Fanuc KAREL source: kt00161.KL

-- PROVISIONAL review KL for V770-1; original PC SHA256 88295595c356cc0f7e4fe96be16e9ae8570dd98f7b765e4e92e81a0925efb0fa
-- Incomplete behavior may be omitted. Consult companion uncertainty JSON. Do not deploy.
PROGRAM KT00161
%NOLOCKGROUP
VAR
  I1 : INTEGER
  I2 : INTEGER
  OUT : INTEGER
BEGIN
  -- UNRESOLVED_PC offsets 5-16; opcodes 2E,23
  -- UNRESOLVED_PC offsets 21-32; opcodes 2E,23
  -- UNRESOLVED_PC offsets 37-48; opcodes 2E,23
  -- UNRESOLVED_PC offsets 53-64; opcodes 2E,23
  -- UNRESOLVED_PC offsets 69-88; opcodes 21,21,56,23
  -- UNRESOLVED_PC offsets 93-97; opcodes 7F
END KT00161
